(* IEC 61131-3 sources: OpenPlc_Lezioni/ST/SR_TIMER1_ST/build, 2 files *)

(* ---- plc.st ---- *)
TYPE
  LOGLEVEL : (CRITICAL, WARNING, INFO, DEBUG) := INFO;
END_TYPE

FUNCTION_BLOCK LOGGER
  VAR_INPUT
    TRIG : BOOL;
    MSG : STRING;
    LEVEL : LOGLEVEL := INFO;
  END_VAR
  VAR
    TRIG0 : BOOL;
  END_VAR

  IF TRIG AND NOT TRIG0 THEN
  {{
   LogMessage(GetFbVar(LEVEL),(char*)GetFbVar(MSG, .body),GetFbVar(MSG, .len));
  }}
  END_IF;
  TRIG0:=TRIG;
END_FUNCTION_BLOCK

PROGRAM program0
  VAR
    bt1 : BOOL;
    bt2 : BOOL;
    led : BOOL;
    timer_ok : BOOL;
    tmer1 : TON;
    sr1 : SR;
  END_VAR

  tmer1(
      IN := bt1,
      PT := T#5s,
      Q => timer_ok
  );

  sr1(
      S1 := timer_ok,
      R := bt2,
      Q1 => led
  );
END_PROGRAM

CONFIGURATION Config0

  RESOURCE Res0 ON PLC
    TASK task0(INTERVAL := T#20ms,PRIORITY := 0);
    PROGRAM instance0 WITH task0 : program0;
  END_RESOURCE
END_CONFIGURATION

(* ---- generated_plc.st ---- *)
PROGRAM program0
  VAR
    bt1 : BOOL;
    bt2 : BOOL;
    led : BOOL;
    timer_ok : BOOL;
    tmer1 : TON;
    sr1 : SR;
  END_VAR

  tmer1(
      IN := bt1,
      PT := T#5s,
      Q => timer_ok
  );

  sr1(
      S1 := timer_ok,
      R := bt2,
      Q1 => led
  );
END_PROGRAM

CONFIGURATION Config0

  RESOURCE Res0 ON PLC
    TASK task0(INTERVAL := T#20ms,PRIORITY := 0);
    PROGRAM instance0 WITH task0 : program0;
  END_RESOURCE
END_CONFIGURATION
